// TIA Portal V20 export
ORGANIZATION_BLOCK "T6_Ciclo"   // OB129, LAD, ProgramCycle
TITLE = T6_Ciclo
{ S7_Optimized_Access := 'TRUE' }
AUTHOR : IA
FAMILY : PRUEBA
VERSION : 0.1
// Tanda 2: llama a todas las pruebas
// stored: AutoNumber false, IsIECCheckEnabled false, SetENOAutomatically false
   VAR_INPUT
      Initial_Call : Bool;
      Remanence : Bool;
   END_VAR
BEGIN

REGION Network 1: T6_S_Base
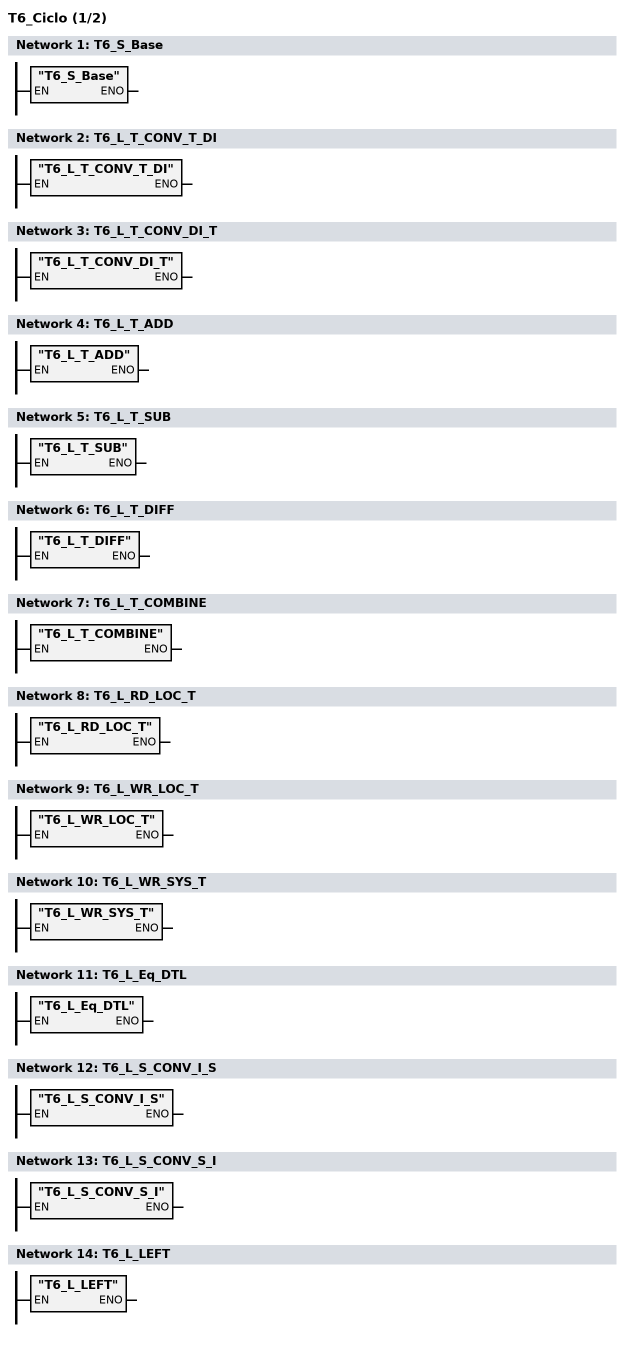
   RUNG wire#powerrail
      "T6_S_Base"()
   END_RUNG
   // the same network as SCL:
   "T6_S_Base"();
END_REGION

REGION Network 2: T6_L_T_CONV_T_DI
   RUNG wire#powerrail
      "T6_L_T_CONV_T_DI"()
   END_RUNG
   // the same network as SCL:
   "T6_L_T_CONV_T_DI"();
END_REGION

REGION Network 3: T6_L_T_CONV_DI_T
   RUNG wire#powerrail
      "T6_L_T_CONV_DI_T"()
   END_RUNG
   // the same network as SCL:
   "T6_L_T_CONV_DI_T"();
END_REGION

REGION Network 4: T6_L_T_ADD
   RUNG wire#powerrail
      "T6_L_T_ADD"()
   END_RUNG
   // the same network as SCL:
   "T6_L_T_ADD"();
END_REGION

REGION Network 5: T6_L_T_SUB
   RUNG wire#powerrail
      "T6_L_T_SUB"()
   END_RUNG
   // the same network as SCL:
   "T6_L_T_SUB"();
END_REGION

REGION Network 6: T6_L_T_DIFF
   RUNG wire#powerrail
      "T6_L_T_DIFF"()
   END_RUNG
   // the same network as SCL:
   "T6_L_T_DIFF"();
END_REGION

REGION Network 7: T6_L_T_COMBINE
   RUNG wire#powerrail
      "T6_L_T_COMBINE"()
   END_RUNG
   // the same network as SCL:
   "T6_L_T_COMBINE"();
END_REGION

REGION Network 8: T6_L_RD_LOC_T
   RUNG wire#powerrail
      "T6_L_RD_LOC_T"()
   END_RUNG
   // the same network as SCL:
   "T6_L_RD_LOC_T"();
END_REGION

REGION Network 9: T6_L_WR_LOC_T
   RUNG wire#powerrail
      "T6_L_WR_LOC_T"()
   END_RUNG
   // the same network as SCL:
   "T6_L_WR_LOC_T"();
END_REGION

REGION Network 10: T6_L_WR_SYS_T
   RUNG wire#powerrail
      "T6_L_WR_SYS_T"()
   END_RUNG
   // the same network as SCL:
   "T6_L_WR_SYS_T"();
END_REGION

REGION Network 11: T6_L_Eq_DTL
   RUNG wire#powerrail
      "T6_L_Eq_DTL"()
   END_RUNG
   // the same network as SCL:
   "T6_L_Eq_DTL"();
END_REGION

REGION Network 12: T6_L_S_CONV_I_S
   RUNG wire#powerrail
      "T6_L_S_CONV_I_S"()
   END_RUNG
   // the same network as SCL:
   "T6_L_S_CONV_I_S"();
END_REGION

REGION Network 13: T6_L_S_CONV_S_I
   RUNG wire#powerrail
      "T6_L_S_CONV_S_I"()
   END_RUNG
   // the same network as SCL:
   "T6_L_S_CONV_S_I"();
END_REGION

REGION Network 14: T6_L_LEFT
   RUNG wire#powerrail
      "T6_L_LEFT"()
   END_RUNG
   // the same network as SCL:
   "T6_L_LEFT"();
END_REGION

REGION Network 15: T6_L_RIGHT
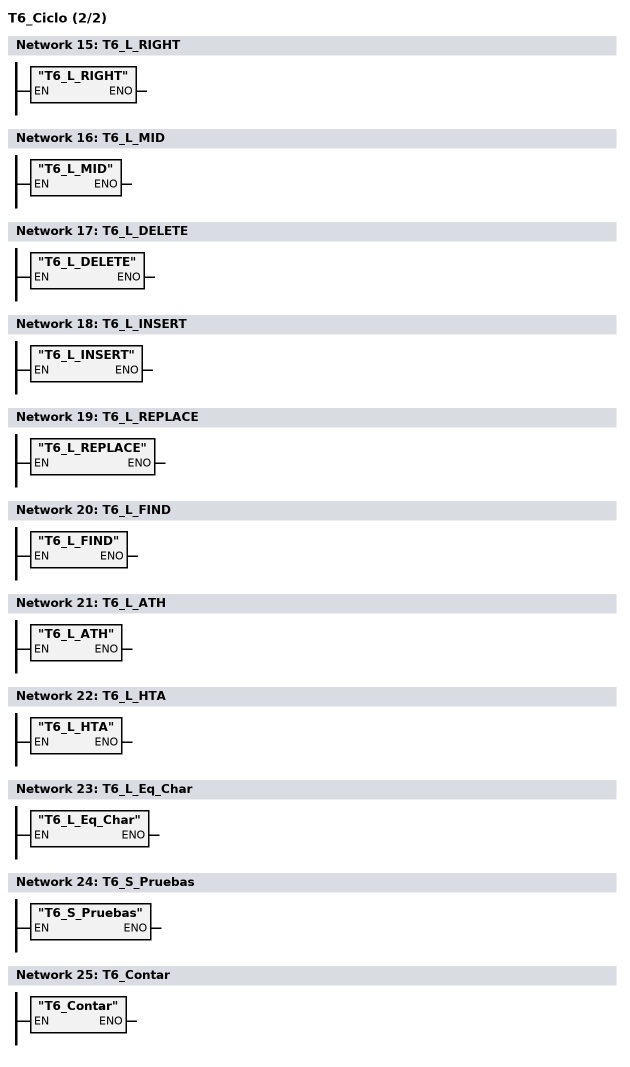
   RUNG wire#powerrail
      "T6_L_RIGHT"()
   END_RUNG
   // the same network as SCL:
   "T6_L_RIGHT"();
END_REGION

REGION Network 16: T6_L_MID
   RUNG wire#powerrail
      "T6_L_MID"()
   END_RUNG
   // the same network as SCL:
   "T6_L_MID"();
END_REGION

REGION Network 17: T6_L_DELETE
   RUNG wire#powerrail
      "T6_L_DELETE"()
   END_RUNG
   // the same network as SCL:
   "T6_L_DELETE"();
END_REGION

REGION Network 18: T6_L_INSERT
   RUNG wire#powerrail
      "T6_L_INSERT"()
   END_RUNG
   // the same network as SCL:
   "T6_L_INSERT"();
END_REGION

REGION Network 19: T6_L_REPLACE
   RUNG wire#powerrail
      "T6_L_REPLACE"()
   END_RUNG
   // the same network as SCL:
   "T6_L_REPLACE"();
END_REGION

REGION Network 20: T6_L_FIND
   RUNG wire#powerrail
      "T6_L_FIND"()
   END_RUNG
   // the same network as SCL:
   "T6_L_FIND"();
END_REGION

REGION Network 21: T6_L_ATH
   RUNG wire#powerrail
      "T6_L_ATH"()
   END_RUNG
   // the same network as SCL:
   "T6_L_ATH"();
END_REGION

REGION Network 22: T6_L_HTA
   RUNG wire#powerrail
      "T6_L_HTA"()
   END_RUNG
   // the same network as SCL:
   "T6_L_HTA"();
END_REGION

REGION Network 23: T6_L_Eq_Char
   RUNG wire#powerrail
      "T6_L_Eq_Char"()
   END_RUNG
   // the same network as SCL:
   "T6_L_Eq_Char"();
END_REGION

REGION Network 24: T6_S_Pruebas
   RUNG wire#powerrail
      "T6_S_Pruebas"()
   END_RUNG
   // the same network as SCL:
   "T6_S_Pruebas"();
END_REGION

REGION Network 25: T6_Contar
   RUNG wire#powerrail
      "T6_Contar"()
   END_RUNG
   // the same network as SCL:
   "T6_Contar"();
END_REGION
END_ORGANIZATION_BLOCK
